(* IEC 61131-3 sources: rk/stdlib/generated, 8 files *)

(* ---- wasi-cli-types.st ---- *)
/* Generated from the WIT of wasi:cli@0.3.0. DO NOT EDIT! */
NAMESPACE INTERNAL Wasi
	NAMESPACE Cli
		NAMESPACE Types
			TYPE ERROR_CODE : USINT (
				IO := 0,
				ILLEGAL_BYTE_SEQUENCE := 1,
				PIPE := 2
			); END_TYPE
		END_NAMESPACE
	END_NAMESPACE
END_NAMESPACE

(* ---- wasi-clocks-system-clock.st ---- *)
/* Generated from the WIT of wasi:clocks@0.3.0. DO NOT EDIT! */
NAMESPACE INTERNAL Wasi
	NAMESPACE Clocks
		/* WASI System Clock is a clock API intended to let users query the current
		   time. The clock is not necessarily monotonic as it may be reset.

		   It is intended to be portable at least between Unix-family platforms and
		   Windows.

		   External references may be reset, so this clock is not necessarily
		   monotonic, making it unsuitable for measuring elapsed time.

		   It is intended for reporting the current date and time for humans. */
		NAMESPACE SystemClock
			/* An "instant", or "exact time", is a point in time without regard to any
			   time zone: just the time since a particular external reference point,
			   often called an "epoch".

			   Here, the epoch is 1970-01-01T00:00:00Z, also known as
			   [POSIX's Seconds Since the Epoch], also known as [Unix Time].

			   Note that even if the seconds field is negative, incrementing
			   nanoseconds always represents moving forwards in time.
			   For example, `{ -1 seconds, 999999999 nanoseconds }` represents the
			   instant one nanosecond before the epoch.
			   For more on various different ways to represent time, see
			   https://tc39.es/proposal-temporal/docs/timezone.html

			   [POSIX's Seconds Since the Epoch]: https://pubs.opengroup.org/onlinepubs/9699919799/xrat/V4_xbd_chap04.html#tag_21_04_16
			   [Unix Time]: https://en.wikipedia.org/wiki/Unix_time */
			TYPE INSTANT : STRUCT
				seconds : LINT;
				nanoseconds : UDINT;
			END_STRUCT END_TYPE

			/* `now` as the host gives it: the values of its result, which `NOW` puts
			   in its members. */
			{extern 'wasi:clocks/system-clock@0.3.0' 'now'}
			FUNCTION PRIVATE NOW_RAW
			VAR_OUTPUT
				seconds : LINT;
				nanoseconds : UDINT;
			END_VAR
			END_FUNCTION

			/* Read the current value of the clock.

			   This clock is not monotonic, therefore calling this function repeatedly
			   will not necessarily produce a sequence of non-decreasing values.

			   The nanoseconds field of the output is always less than 1000000000. */
			FUNCTION NOW : INSTANT
				NOW_RAW(seconds => NOW.seconds, nanoseconds => NOW.nanoseconds);
			END_FUNCTION

			/* Query the resolution of the clock. Returns the smallest duration of time
			   that the implementation permits distinguishing. */
			{extern 'wasi:clocks/system-clock@0.3.0' 'get-resolution'}
			FUNCTION GET_RESOLUTION : Wasi.Clocks.Types.DURATION
			END_FUNCTION
		END_NAMESPACE
	END_NAMESPACE
END_NAMESPACE

(* ---- wasi-clocks-types.st ---- *)
/* Generated from the WIT of wasi:clocks@0.3.0. DO NOT EDIT! */
NAMESPACE INTERNAL Wasi
	NAMESPACE Clocks
		/* This interface common types used throughout wasi:clocks. */
		NAMESPACE Types
			/* A duration of time, in nanoseconds. */
			TYPE DURATION : ULINT; END_TYPE
		END_NAMESPACE
	END_NAMESPACE
END_NAMESPACE

(* ---- wasi-clocks-timezone.st ---- *)
/* Generated from the WIT of wasi:clocks@0.3.0. DO NOT EDIT! */
NAMESPACE INTERNAL Wasi
	NAMESPACE Clocks
		NAMESPACE Timezone
			/* `iana-id` as the host gives it: its result in words of 8 bytes, as the
			   canonical ABI lays it out, which `IANA_ID` reads, and its string in
			   `value`, where the host writes it. */
			{extern 'wasi:clocks/timezone@0.3.0' 'iana-id'}
			FUNCTION PRIVATE IANA_ID_RAW
			VAR_IN_OUT
				value : STRING;
			END_VAR
			VAR_OUTPUT
				w0 : LWORD;
				w1 : LWORD;
			END_VAR
			END_FUNCTION

			/* Return the IANA identifier of the currently configured timezone. This
			   should be an identifier from the IANA Time Zone Database.

			   For displaying to a user, the identifier should be converted into a
			   localized name by means of an internationalization API.

			   If the implementation does not expose an actual timezone, or is unable
			   to provide mappings from times to deltas between the configured timezone
			   and UTC, or determining the current timezone fails, or the timezone does
			   not have an IANA identifier, this returns nothing. */
			FUNCTION IANA_ID
			VAR_IN_OUT
				value : STRING;
			END_VAR
			VAR_OUTPUT
				is_some : BOOL;
			END_VAR
			VAR
				w0 : LWORD;
				w1 : LWORD;
			END_VAR
				IANA_ID_RAW(value := value, w0 => w0, w1 => w1);
				is_some := w0.%X0;
			END_FUNCTION

			/* `utc-offset` as the host takes it: its parameters as the canonical ABI
			   passes them, which `UTC_OFFSET` passes field by field. */
			{extern 'wasi:clocks/timezone@0.3.0' 'utc-offset'}
			FUNCTION PRIVATE UTC_OFFSET_RAW
			VAR_INPUT
				when_seconds : LINT;
				when_nanoseconds : UDINT;
			END_VAR
			VAR_OUTPUT
				is_some : BOOL;
				value : LINT;
			END_VAR
			END_FUNCTION

			/* The number of nanoseconds difference between UTC time and the local
			   time of the currently configured timezone, at the exact time of
			   `instant`.

			   The magnitude of the returned value will always be less than
			   86,400,000,000,000 which is the number of nanoseconds in a day
			   (24*60*60*1e9).

			   If the implementation does not expose an actual timezone, or is unable
			   to provide mappings from times to deltas between the configured timezone
			   and UTC, or determining the current timezone fails, this returns
			   nothing. */
			FUNCTION UTC_OFFSET
			VAR_INPUT
				when : Wasi.Clocks.SystemClock.INSTANT;
			END_VAR
			VAR_OUTPUT
				is_some : BOOL;
				value : LINT;
			END_VAR
				UTC_OFFSET_RAW(when_seconds := when.seconds, when_nanoseconds := when.nanoseconds, is_some => is_some, value => value);
			END_FUNCTION

			/* `to-debug-string` as the host gives it: its result in words of 8 bytes,
			   as the canonical ABI lays it out, which `TO_DEBUG_STRING` reads, and its
			   string in `value`, where the host writes it. */
			{extern 'wasi:clocks/timezone@0.3.0' 'to-debug-string'}
			FUNCTION PRIVATE TO_DEBUG_STRING_RAW
			VAR_IN_OUT
				value : STRING;
			END_VAR
			VAR_OUTPUT
				w0 : LWORD;
				w1 : LWORD;
			END_VAR
			END_FUNCTION

			/* Returns a string that is suitable to assist humans in debugging whether
			   any timezone is available, and if so, which. This may be the same string
			   as `iana-id`, or a formatted representation of the UTC offset such as
			   `-04:00`, or something else.

			   WARNING: The returned string should not be consumed mechanically! It may
			   change across platforms, hosts, or other implementation details. Parsing
			   this string is a major platform-compatibility hazard. */
			FUNCTION TO_DEBUG_STRING
			VAR_IN_OUT
				value : STRING;
			END_VAR
			VAR
				w0 : LWORD;
				w1 : LWORD;
			END_VAR
				TO_DEBUG_STRING_RAW(value := value, w0 => w0, w1 => w1);
			END_FUNCTION
		END_NAMESPACE
	END_NAMESPACE
END_NAMESPACE

(* ---- wasi-cli-stderr.st ---- *)
/* Generated from the WIT of wasi:cli@0.3.0. DO NOT EDIT! */
NAMESPACE INTERNAL Wasi
	NAMESPACE Cli
		NAMESPACE Stderr
			/* Write the given stream to stderr.

			   If the stream's writable end is dropped this function will either return
			   success once the entire contents of the stream have been written or an
			   error-code representing a failure.

			   Otherwise if there is an error the readable end of the stream will be
			   dropped and this function will return an error-code. */
			{extern 'wasi:cli/stderr@0.3.0' 'write-via-stream'}
			FUNCTION WRITE_VIA_STREAM : UDINT
			VAR_INPUT
				data : UDINT;
			END_VAR
			END_FUNCTION

			/* Makes a stream of `u8`, and gives its reading end, then its writing end. */
			{extern 'wasi:cli/stderr@0.3.0' '[stream-new-0]write-via-stream'}
			FUNCTION BYTES_STREAM_NEW
			VAR_OUTPUT
				readable : UDINT;
				writable : UDINT;
			END_VAR
			END_FUNCTION

			/* Writes the bytes of `data`, as many as the reader takes: `written` of
			   them, after `DONE`. `closed` is TRUE once the reader has let go. */
			{extern async 'wasi:cli/stderr@0.3.0' '[stream-write-0]write-via-stream'}
			FUNCTION_BLOCK BYTES_STREAM_WRITE
			VAR_INPUT
				stream : UDINT;
				data : STRING[4096];
			END_VAR
			VAR_OUTPUT
				DONE : BOOL;
				written : UDINT;
				closed : BOOL;
			END_VAR
			END_FUNCTION_BLOCK

			/* Writes the `count` bytes from the one `data` points at, as many as the
			   reader takes: `written` of them, after `DONE`. The host reads them where
			   they are while the write runs, so they stay there, unchanged, until
			   `DONE`. `closed` is TRUE once the reader has let go. */
			{extern async 'wasi:cli/stderr@0.3.0' '[stream-write-0]write-via-stream'}
			FUNCTION_BLOCK BYTES_STREAM_WRITE_ARRAY
			VAR_INPUT
				stream : UDINT;
				data : REF_TO BYTE;
				count : UDINT;
			END_VAR
			VAR_OUTPUT
				DONE : BOOL;
				written : UDINT;
				closed : BOOL;
			END_VAR
			END_FUNCTION_BLOCK

			/* Lets go of the stream's reading end, `stream`. */
			{extern 'wasi:cli/stderr@0.3.0' '[stream-drop-readable-0]write-via-stream'}
			FUNCTION BYTES_STREAM_DROP_READABLE
			VAR_INPUT
				stream : UDINT;
			END_VAR
			END_FUNCTION

			/* Lets go of the stream's writing end, `stream`. */
			{extern 'wasi:cli/stderr@0.3.0' '[stream-drop-writable-0]write-via-stream'}
			FUNCTION BYTES_STREAM_DROP_WRITABLE
			VAR_INPUT
				stream : UDINT;
			END_VAR
			END_FUNCTION

			/* The bytes `IN` holds, which `BYTES_STREAM_WRITER` counts. */
			FUNCTION PRIVATE BYTES_STREAM_TEXT_LEN : UDINT
			VAR_INPUT
				IN : STRING[4096];
			END_VAR
				{wasm 'str.byte_len' (params IN) (result BYTES_STREAM_TEXT_LEN)}
			END_FUNCTION

			/* `IN` without its first `L` bytes: what `BYTES_STREAM_WRITER` has left to
			   write. */
			FUNCTION PRIVATE BYTES_STREAM_TEXT_AFTER : STRING[4096]
			VAR_INPUT
				IN : STRING[4096];
				L : UDINT;
			END_VAR
			VAR
				P : UDINT := 1;
			END_VAR
				{wasm 'str.byte_delete' (params IN L P) (result BYTES_STREAM_TEXT_AFTER)}
			END_FUNCTION

			/* Writes text to a stream of bytes it makes at its first call, for the
			   function `readable` is handed to. */
			FUNCTION_BLOCK BYTES_STREAM_WRITER
			VAR_INPUT
				/* A rising edge writes `IN`. An edge while `BUSY` is ignored. */
				REQ : BOOL;
				/* The text to write. */
				IN : STRING[4096];
				/* A rising edge ends the stream, once no write is under way. */
				CLOSE : BOOL;
			END_VAR
			VAR_OUTPUT
				/* The stream's reading end, to hand to the function that reads it. */
				readable : UDINT;
				/* TRUE while the reader has not taken all of `IN`. */
				BUSY : BOOL;
				/* TRUE in the call where the reader has taken all of `IN`, at once for an
				   empty text. */
				DONE : BOOL;
				/* TRUE once a write finds the reader gone, or a request comes after
				   `CLOSE`: the stream does not open again. */
				ERROR : BOOL;
			END_VAR
			VAR
				writable : UDINT;
				requested : BOOL;
				closing : BOOL;
				shut : BOOL;
				closed : BOOL;
				rest : STRING[4096];
				write : BYTES_STREAM_WRITE;
			END_VAR
			VAR_TEMP
				again : BOOL;
			END_VAR
				IF writable = 0 AND NOT closed THEN
					BYTES_STREAM_NEW(readable => readable, writable => writable);
				END_IF;
				DONE := FALSE;
				// An edge while BUSY is ignored.
				IF REQ AND NOT requested AND NOT BUSY THEN
					ERROR := closed;
					IF NOT closed THEN
						// A write of no bytes asks the reader whether it is ready,
						// which it may answer late: an empty text is done here.
						IF BYTES_STREAM_TEXT_LEN(IN) = 0 THEN
							DONE := TRUE;
						ELSE
							rest := IN;
							BUSY := TRUE;
						END_IF;
					END_IF;
				END_IF;
				requested := REQ;
				IF BUSY THEN
					// Each pass after the first hands over a byte at least, so the
					// loop ends.
					REPEAT
						again := FALSE;
						// Starts the write of the rest, or checks the one running.
						write(stream := writable, data := rest);
						IF write.DONE THEN
							IF write.closed THEN
								// The reader left: the writing end goes too.
								BYTES_STREAM_DROP_WRITABLE(stream := writable);
								writable := 0;
								closed := TRUE;
								BUSY := FALSE;
								ERROR := TRUE;
							ELSIF write.written < BYTES_STREAM_TEXT_LEN(rest) THEN
								// The reader took a part: the rest goes next, at once while
								// it takes some.
								rest := BYTES_STREAM_TEXT_AFTER(rest, write.written);
								again := write.written > 0;
							ELSE
								BUSY := FALSE;
								DONE := TRUE;
							END_IF;
						END_IF;
					UNTIL NOT again
					END_REPEAT;
				END_IF;
				// The writing end goes once no write is under way.
				IF CLOSE AND NOT closing THEN
					shut := TRUE;
				END_IF;
				closing := CLOSE;
				IF shut AND NOT BUSY THEN
					IF writable <> 0 THEN
						BYTES_STREAM_DROP_WRITABLE(stream := writable);
						writable := 0;
					END_IF;
					closed := TRUE;
					shut := FALSE;
				END_IF;
			END_FUNCTION_BLOCK

			/* The subscript of the first byte of `IN`, which
			   `BYTES_STREAM_ARRAY_WRITER` writes from. */
			FUNCTION PRIVATE BYTES_STREAM_ARRAY_FIRST : LINT
			VAR_INPUT
				IN : ARRAY[*] OF BYTE;
			END_VAR
			VAR
				DIM : DINT := 1;
			END_VAR
				{wasm 'array.lower_bound' (params IN DIM) (result BYTES_STREAM_ARRAY_FIRST)}
			END_FUNCTION

			/* How many bytes `IN` holds, which `BYTES_STREAM_ARRAY_WRITER` writes at
			   most. */
			FUNCTION PRIVATE BYTES_STREAM_ARRAY_LEN : LINT
			VAR_INPUT
				IN : ARRAY[*] OF BYTE;
			END_VAR
			VAR
				DIM : DINT := 1;
				lower : LINT;
				upper : LINT;
			END_VAR
				{wasm 'array.lower_bound' (params IN DIM) (result lower)}
				{wasm 'array.upper_bound' (params IN DIM) (result upper)}
				BYTES_STREAM_ARRAY_LEN := upper - lower + 1;
			END_FUNCTION

			/* Writes bytes from an array to a stream of bytes it makes at its first
			   call, for the function `readable` is handed to. */
			FUNCTION_BLOCK BYTES_STREAM_ARRAY_WRITER
			VAR_INPUT
				/* A rising edge writes the first `COUNT` bytes of `IN`. An edge while
				   `BUSY` is ignored. */
				REQ : BOOL;
				/* How many bytes of `IN` a request writes, from its first on. */
				COUNT : UDINT;
				/* A rising edge ends the stream, once no write is under way. */
				CLOSE : BOOL;
			END_VAR
			VAR_IN_OUT
				/* The bytes to write. The host reads them where they are while `BUSY`:
				   they stay as they are until `DONE`. */
				IN : ARRAY[*] OF BYTE;
			END_VAR
			VAR_OUTPUT
				/* The stream's reading end, to hand to the function that reads it. */
				readable : UDINT;
				/* TRUE while the reader has not taken all `COUNT` bytes. */
				BUSY : BOOL;
				/* TRUE in the call where the reader has taken all `COUNT` bytes, at once
				   for none. */
				DONE : BOOL;
				/* TRUE once a write finds the reader gone, or a request comes after
				   `CLOSE`: the stream does not open again. */
				ERROR : BOOL;
			END_VAR
			VAR
				writable : UDINT;
				requested : BOOL;
				closing : BOOL;
				shut : BOOL;
				closed : BOOL;
				total : UDINT;
				sent : UDINT;
				base : LINT;
				write : BYTES_STREAM_WRITE_ARRAY;
			END_VAR
			VAR_TEMP
				again : BOOL;
				offset : LINT;
			END_VAR
				IF writable = 0 AND NOT closed THEN
					BYTES_STREAM_NEW(readable => readable, writable => writable);
				END_IF;
				DONE := FALSE;
				// An edge while BUSY is ignored.
				IF REQ AND NOT requested AND NOT BUSY THEN
					ERROR := closed;
					IF NOT closed THEN
						// A write of no bytes asks the reader whether it is ready,
						// which it may answer late: none is done here.
						IF COUNT = 0 THEN
							DONE := TRUE;
						ELSIF COUNT > BYTES_STREAM_ARRAY_LEN(IN) THEN
							__RAISE('COUNT is past the end of IN');
						ELSE
							total := COUNT;
							sent := 0;
							base := BYTES_STREAM_ARRAY_FIRST(IN);
							BUSY := TRUE;
						END_IF;
					END_IF;
				END_IF;
				requested := REQ;
				IF BUSY THEN
					// Each pass after the first hands over a byte at least, so the
					// loop ends.
					REPEAT
						again := FALSE;
						offset := sent;
						// Starts the write of the bytes not taken yet, from where they
						// are, or checks the one running.
						write(stream := writable, data := REF(IN[base + offset]), count := total - sent);
						IF write.DONE THEN
							IF write.closed THEN
								// The reader left: the writing end goes too.
								BYTES_STREAM_DROP_WRITABLE(stream := writable);
								writable := 0;
								closed := TRUE;
								BUSY := FALSE;
								ERROR := TRUE;
							ELSIF write.written < total - sent THEN
								// The reader took a part: the rest goes next, at once while
								// it takes some.
								sent := sent + write.written;
								again := write.written > 0;
							ELSE
								BUSY := FALSE;
								DONE := TRUE;
							END_IF;
						END_IF;
					UNTIL NOT again
					END_REPEAT;
				END_IF;
				// The writing end goes once no write is under way.
				IF CLOSE AND NOT closing THEN
					shut := TRUE;
				END_IF;
				closing := CLOSE;
				IF shut AND NOT BUSY THEN
					IF writable <> 0 THEN
						BYTES_STREAM_DROP_WRITABLE(stream := writable);
						writable := 0;
					END_IF;
					closed := TRUE;
					shut := FALSE;
				END_IF;
			END_FUNCTION_BLOCK

			/* Reads the value the future holds, which comes back after `DONE`. */
			{extern async 'wasi:cli/stderr@0.3.0' '[future-read-1]write-via-stream'}
			FUNCTION_BLOCK RESULT_FUTURE_READ
			VAR_INPUT
				future : UDINT;
			END_VAR
			VAR_OUTPUT
				DONE : BOOL;
				failed : BOOL;
				error : Wasi.Cli.Types.ERROR_CODE;
			END_VAR
			END_FUNCTION_BLOCK

			/* Lets go of the future's reading end, `future`. */
			{extern 'wasi:cli/stderr@0.3.0' '[future-drop-readable-1]write-via-stream'}
			FUNCTION RESULT_FUTURE_DROP_READABLE
			VAR_INPUT
				future : UDINT;
			END_VAR
			END_FUNCTION

			/* Reads the value the future holds, which comes back after `DONE`, then
			   lets go of the future's reading end: `future` is 0 from then on, and a
			   call with `future` 0 does nothing. */
			FUNCTION_BLOCK RESULT_FUTURE_GET
			VAR_IN_OUT
				future : UDINT;
			END_VAR
			VAR_OUTPUT
				DONE : BOOL;
				failed : BOOL;
				error : Wasi.Cli.Types.ERROR_CODE;
			END_VAR
			VAR
				call : RESULT_FUTURE_READ;
			END_VAR
				DONE := FALSE;
				IF future <> 0 THEN
					call(future := future);
					IF call.DONE THEN
						failed := call.failed;
						error := call.error;
						RESULT_FUTURE_DROP_READABLE(future := future);
						future := 0;
						DONE := TRUE;
					END_IF;
				END_IF;
			END_FUNCTION_BLOCK

			/* Writes text to `write-via-stream` through a stream of bytes it opens at
			   the first request. */
			FUNCTION_BLOCK WRITE_VIA_STREAM_WRITER
			VAR_INPUT
				/* A rising edge writes `IN`; the first opens the stream and calls
				   `write-via-stream` with it. An edge while `BUSY` is ignored. */
				REQ : BOOL;
				/* The text to write. */
				IN : STRING[4096];
				/* A rising edge ends the stream, once no write is under way. */
				CLOSE : BOOL;
			END_VAR
			VAR_OUTPUT
				/* TRUE while the reader has not taken all of `IN`. */
				BUSY : BOOL;
				/* TRUE in the call where the reader has taken all of `IN`, at once for an
				   empty text. */
				DONE : BOOL;
				/* TRUE once a write finds the reader gone, a request comes after `CLOSE`,
				   or the `result<_, error-code>` from `write-via-stream` is an error,
				   whose `error-code` is in `ERRORID`. */
				ERROR : BOOL;
				/* The `error-code` of the `result<_, error-code>` from `write-via-stream`,
				   when it is an error, which turns `ERROR` TRUE. */
				ERRORID : Wasi.Cli.Types.ERROR_CODE;
				/* TRUE once the `future<result<_, error-code>>` from `write-via-stream`
				   has its value. */
				ENDED : BOOL;
			END_VAR
			VAR
				open : BOOL;
				stream : BYTES_STREAM_WRITER;
				future : UDINT;
				answer : RESULT_FUTURE_GET;
			END_VAR
				// The stream, made at the first request and handed to the function.
				IF REQ AND NOT open THEN
					stream(REQ := FALSE, IN := IN, CLOSE := FALSE);
					future := Wasi.Cli.Stderr.WRITE_VIA_STREAM(data := stream.readable);
					open := TRUE;
				END_IF;
				IF open THEN
					stream(REQ := REQ, IN := IN, CLOSE := CLOSE);
					BUSY := stream.BUSY;
					DONE := stream.DONE;
					// The answer, read once it comes, and kept.
					answer(future := future);
					IF answer.DONE THEN
						ERRORID := answer.error;
						ENDED := TRUE;
					END_IF;
					ERROR := stream.ERROR OR answer.failed;
				END_IF;
			END_FUNCTION_BLOCK

			/* Writes bytes from an array to `write-via-stream` through a stream of
			   bytes it opens at the first request. */
			FUNCTION_BLOCK WRITE_VIA_STREAM_ARRAY_WRITER
			VAR_INPUT
				/* A rising edge writes the first `COUNT` bytes of `IN`; the first opens
				   the stream and calls `write-via-stream` with it. An edge while `BUSY` is
				   ignored. */
				REQ : BOOL;
				/* How many bytes of `IN` a request writes, from its first on. */
				COUNT : UDINT;
				/* A rising edge ends the stream, once no write is under way. */
				CLOSE : BOOL;
			END_VAR
			VAR_IN_OUT
				/* The bytes to write. The host reads them where they are while `BUSY`:
				   they stay as they are until `DONE`. */
				IN : ARRAY[*] OF BYTE;
			END_VAR
			VAR_OUTPUT
				/* TRUE while the reader has not taken all `COUNT` bytes. */
				BUSY : BOOL;
				/* TRUE in the call where the reader has taken all `COUNT` bytes, at once
				   for none. */
				DONE : BOOL;
				/* TRUE once a write finds the reader gone, a request comes after `CLOSE`,
				   or the `result<_, error-code>` from `write-via-stream` is an error,
				   whose `error-code` is in `ERRORID`. */
				ERROR : BOOL;
				/* The `error-code` of the `result<_, error-code>` from `write-via-stream`,
				   when it is an error, which turns `ERROR` TRUE. */
				ERRORID : Wasi.Cli.Types.ERROR_CODE;
				/* TRUE once the `future<result<_, error-code>>` from `write-via-stream`
				   has its value. */
				ENDED : BOOL;
			END_VAR
			VAR
				open : BOOL;
				stream : BYTES_STREAM_ARRAY_WRITER;
				future : UDINT;
				answer : RESULT_FUTURE_GET;
			END_VAR
				// The stream, made at the first request and handed to the function.
				IF REQ AND NOT open THEN
					stream(REQ := FALSE, COUNT := COUNT, CLOSE := FALSE, IN := IN);
					future := Wasi.Cli.Stderr.WRITE_VIA_STREAM(data := stream.readable);
					open := TRUE;
				END_IF;
				IF open THEN
					stream(REQ := REQ, COUNT := COUNT, CLOSE := CLOSE, IN := IN);
					BUSY := stream.BUSY;
					DONE := stream.DONE;
					// The answer, read once it comes, and kept.
					answer(future := future);
					IF answer.DONE THEN
						ERRORID := answer.error;
						ENDED := TRUE;
					END_IF;
					ERROR := stream.ERROR OR answer.failed;
				END_IF;
			END_FUNCTION_BLOCK
		END_NAMESPACE
	END_NAMESPACE
END_NAMESPACE
/* Not generated:
   - `BYTES_STREAM_CANCEL_WRITE`: a cancel blocks the scan.
   - `RESULT_FUTURE_CANCEL_READ`: a cancel blocks the scan. */

(* ---- wasi-cli-stdin.st ---- *)
/* Generated from the WIT of wasi:cli@0.3.0. DO NOT EDIT! */
NAMESPACE INTERNAL Wasi
	NAMESPACE Cli
		NAMESPACE Stdin
			/* Return a stream for reading from stdin.

			   This function returns a stream which provides data read from stdin,
			   and a future to signal read results.

			   If the stream's readable end is dropped the future will resolve to success.

			   If the stream's writable end is dropped the future will either resolve to
			   success if stdin was closed by the writer or to an error-code if reading
			   failed for some other reason.

			   Multiple streams may be active at the same time. The behavior of concurrent
			   reads is implementation-specific. */
			{extern 'wasi:cli/stdin@0.3.0' 'read-via-stream'}
			FUNCTION READ_VIA_STREAM
			VAR_OUTPUT
				item0 : UDINT;
				item1 : UDINT;
			END_VAR
			END_FUNCTION

			/* Reads the bytes that come next into `data`, as many as it holds at most:
			   `read` of them, after `DONE`. `closed` is TRUE once the writer has let
			   go. */
			{extern async 'wasi:cli/stdin@0.3.0' '[stream-read-0]read-via-stream'}
			FUNCTION_BLOCK BYTES_STREAM_READ
			VAR_INPUT
				stream : UDINT;
			END_VAR
			VAR_OUTPUT
				DONE : BOOL;
				data : STRING[4096];
				read : UDINT;
				closed : BOOL;
			END_VAR
			END_FUNCTION_BLOCK

			/* Reads the bytes that come next into `data`, as many as it holds at most:
			   `read` of them, after `DONE`. `closed` is TRUE once the writer has let
			   go. */
			{extern async 'wasi:cli/stdin@0.3.0' '[stream-read-0]read-via-stream'}
			FUNCTION_BLOCK BYTES_STREAM_READ_ARRAY
			VAR_INPUT
				stream : UDINT;
			END_VAR
			VAR_OUTPUT
				DONE : BOOL;
				data : ARRAY[0..8191] OF BYTE;
				read : UDINT;
				closed : BOOL;
			END_VAR
			END_FUNCTION_BLOCK

			/* Lets go of the stream's reading end, `stream`. */
			{extern 'wasi:cli/stdin@0.3.0' '[stream-drop-readable-0]read-via-stream'}
			FUNCTION BYTES_STREAM_DROP_READABLE
			VAR_INPUT
				stream : UDINT;
			END_VAR
			END_FUNCTION

			/* Reads the value the future holds, which comes back after `DONE`. */
			{extern async 'wasi:cli/stdin@0.3.0' '[future-read-1]read-via-stream'}
			FUNCTION_BLOCK RESULT_FUTURE_READ
			VAR_INPUT
				future : UDINT;
			END_VAR
			VAR_OUTPUT
				DONE : BOOL;
				failed : BOOL;
				error : Wasi.Cli.Types.ERROR_CODE;
			END_VAR
			END_FUNCTION_BLOCK

			/* Lets go of the future's reading end, `future`. */
			{extern 'wasi:cli/stdin@0.3.0' '[future-drop-readable-1]read-via-stream'}
			FUNCTION RESULT_FUTURE_DROP_READABLE
			VAR_INPUT
				future : UDINT;
			END_VAR
			END_FUNCTION

			/* Reads the value the future holds, which comes back after `DONE`, then
			   lets go of the future's reading end: `future` is 0 from then on, and a
			   call with `future` 0 does nothing. */
			FUNCTION_BLOCK RESULT_FUTURE_GET
			VAR_IN_OUT
				future : UDINT;
			END_VAR
			VAR_OUTPUT
				DONE : BOOL;
				failed : BOOL;
				error : Wasi.Cli.Types.ERROR_CODE;
			END_VAR
			VAR
				call : RESULT_FUTURE_READ;
			END_VAR
				DONE := FALSE;
				IF future <> 0 THEN
					call(future := future);
					IF call.DONE THEN
						failed := call.failed;
						error := call.error;
						RESULT_FUTURE_DROP_READABLE(future := future);
						future := 0;
						DONE := TRUE;
					END_IF;
				END_IF;
			END_FUNCTION_BLOCK

			/* Reads what `read-via-stream` gives through a stream of bytes, a request
			   at a time. */
			FUNCTION_BLOCK READ_VIA_STREAM_READER
			VAR_INPUT
				/* A rising edge reads what comes next, 4096 bytes at most; the first calls
				   `read-via-stream`. An edge while `BUSY` is ignored, and one after the
				   stream ended is `DONE` at once, `OUT` empty. */
				REQ : BOOL;
				/* A rising edge lets go of the stream, once no read is under way. */
				CLOSE : BOOL;
			END_VAR
			VAR_OUTPUT
				/* TRUE while a read waits for bytes. */
				BUSY : BOOL;
				/* TRUE in the call where a read has given what came, in `OUT`. */
				DONE : BOOL;
				/* What the last read gave: empty once the stream has ended, nothing more
				   coming. */
				OUT : STRING[4096];
				/* TRUE once the `result<_, error-code>` from `read-via-stream` is an
				   error, whose `error-code` is in `ERRORID`. */
				ERROR : BOOL;
				/* The `error-code` of the `result<_, error-code>` from `read-via-stream`,
				   when it is an error, which turns `ERROR` TRUE. */
				ERRORID : Wasi.Cli.Types.ERROR_CODE;
				/* TRUE once the stream has ended and the `future<result<_, error-code>>`
				   from `read-via-stream` has its value. */
				ENDED : BOOL;
			END_VAR
			VAR
				open : BOOL;
				requested : BOOL;
				closing : BOOL;
				shut : BOOL;
				stream : UDINT;
				future : UDINT;
				read : BYTES_STREAM_READ;
				answer : RESULT_FUTURE_GET;
				came : BOOL;
			END_VAR
				DONE := FALSE;
				// The stream, given by the function at the first request.
				IF REQ AND NOT open THEN
					Wasi.Cli.Stdin.READ_VIA_STREAM(item0 => stream, item1 => future);
					open := TRUE;
				END_IF;
				IF open THEN
					// An edge while BUSY is ignored.
					IF REQ AND NOT requested AND NOT BUSY THEN
						IF stream <> 0 THEN
							BUSY := TRUE;
						ELSE
							// The stream has ended: nothing more comes.
							OUT := '';
							DONE := TRUE;
						END_IF;
					END_IF;
					requested := REQ;
					IF BUSY THEN
						// Starts the read, or checks the one running.
						read(stream := stream);
						IF read.DONE THEN
							OUT := read.data;
							BUSY := FALSE;
							DONE := TRUE;
							IF read.closed THEN
								// The writer left: the reading end goes too.
								BYTES_STREAM_DROP_READABLE(stream := stream);
								stream := 0;
							END_IF;
						END_IF;
					END_IF;
					// The reading end goes on CLOSE, once no read is under way.
					IF CLOSE AND NOT closing THEN
						shut := TRUE;
					END_IF;
					closing := CLOSE;
					IF shut AND NOT BUSY THEN
						IF stream <> 0 THEN
							BYTES_STREAM_DROP_READABLE(stream := stream);
							stream := 0;
						END_IF;
						shut := FALSE;
					END_IF;
					// The answer, read once it comes, and kept.
					answer(future := future);
					IF answer.DONE THEN
						ERRORID := answer.error;
						came := TRUE;
					END_IF;
					ENDED := stream = 0 AND came;
					ERROR := answer.failed;
				END_IF;
			END_FUNCTION_BLOCK

			/* Reads what `read-via-stream` gives through a stream of bytes into an
			   array, a request at a time. */
			FUNCTION_BLOCK READ_VIA_STREAM_ARRAY_READER
			VAR_INPUT
				/* A rising edge reads what comes next, 8192 bytes at most; the first calls
				   `read-via-stream`. An edge while `BUSY` is ignored, and one after the
				   stream ended is `DONE` at once, `COUNT` 0. */
				REQ : BOOL;
				/* A rising edge lets go of the stream, once no read is under way. */
				CLOSE : BOOL;
			END_VAR
			VAR_OUTPUT
				/* TRUE while a read waits for bytes. */
				BUSY : BOOL;
				/* TRUE in the call where a read has given what came, in `OUT`. */
				DONE : BOOL;
				/* The bytes the last read gave, its first `COUNT`. */
				OUT : ARRAY[0..8191] OF BYTE;
				/* How many bytes the last read gave: 0 once the stream has ended, nothing
				   more coming. */
				COUNT : UDINT;
				/* TRUE once the `result<_, error-code>` from `read-via-stream` is an
				   error, whose `error-code` is in `ERRORID`. */
				ERROR : BOOL;
				/* The `error-code` of the `result<_, error-code>` from `read-via-stream`,
				   when it is an error, which turns `ERROR` TRUE. */
				ERRORID : Wasi.Cli.Types.ERROR_CODE;
				/* TRUE once the stream has ended and the `future<result<_, error-code>>`
				   from `read-via-stream` has its value. */
				ENDED : BOOL;
			END_VAR
			VAR
				open : BOOL;
				requested : BOOL;
				closing : BOOL;
				shut : BOOL;
				stream : UDINT;
				future : UDINT;
				read : BYTES_STREAM_READ_ARRAY;
				answer : RESULT_FUTURE_GET;
				came : BOOL;
			END_VAR
				DONE := FALSE;
				// The stream, given by the function at the first request.
				IF REQ AND NOT open THEN
					Wasi.Cli.Stdin.READ_VIA_STREAM(item0 => stream, item1 => future);
					open := TRUE;
				END_IF;
				IF open THEN
					// An edge while BUSY is ignored.
					IF REQ AND NOT requested AND NOT BUSY THEN
						IF stream <> 0 THEN
							BUSY := TRUE;
						ELSE
							// The stream has ended: nothing more comes.
							COUNT := 0;
							DONE := TRUE;
						END_IF;
					END_IF;
					requested := REQ;
					IF BUSY THEN
						// Starts the read, or checks the one running.
						read(stream := stream);
						IF read.DONE THEN
							OUT := read.data;
							COUNT := read.read;
							BUSY := FALSE;
							DONE := TRUE;
							IF read.closed THEN
								// The writer left: the reading end goes too.
								BYTES_STREAM_DROP_READABLE(stream := stream);
								stream := 0;
							END_IF;
						END_IF;
					END_IF;
					// The reading end goes on CLOSE, once no read is under way.
					IF CLOSE AND NOT closing THEN
						shut := TRUE;
					END_IF;
					closing := CLOSE;
					IF shut AND NOT BUSY THEN
						IF stream <> 0 THEN
							BYTES_STREAM_DROP_READABLE(stream := stream);
							stream := 0;
						END_IF;
						shut := FALSE;
					END_IF;
					// The answer, read once it comes, and kept.
					answer(future := future);
					IF answer.DONE THEN
						ERRORID := answer.error;
						came := TRUE;
					END_IF;
					ENDED := stream = 0 AND came;
					ERROR := answer.failed;
				END_IF;
			END_FUNCTION_BLOCK
		END_NAMESPACE
	END_NAMESPACE
END_NAMESPACE
/* Not generated:
   - `BYTES_STREAM_CANCEL_READ`: a cancel blocks the scan.
   - `RESULT_FUTURE_CANCEL_READ`: a cancel blocks the scan. */

(* ---- wasi-cli-stdout.st ---- *)
/* Generated from the WIT of wasi:cli@0.3.0. DO NOT EDIT! */
NAMESPACE INTERNAL Wasi
	NAMESPACE Cli
		NAMESPACE Stdout
			/* Write the given stream to stdout.

			   If the stream's writable end is dropped this function will either return
			   success once the entire contents of the stream have been written or an
			   error-code representing a failure.

			   Otherwise if there is an error the readable end of the stream will be
			   dropped and this function will return an error-code. */
			{extern 'wasi:cli/stdout@0.3.0' 'write-via-stream'}
			FUNCTION WRITE_VIA_STREAM : UDINT
			VAR_INPUT
				data : UDINT;
			END_VAR
			END_FUNCTION

			/* Makes a stream of `u8`, and gives its reading end, then its writing end. */
			{extern 'wasi:cli/stdout@0.3.0' '[stream-new-0]write-via-stream'}
			FUNCTION BYTES_STREAM_NEW
			VAR_OUTPUT
				readable : UDINT;
				writable : UDINT;
			END_VAR
			END_FUNCTION

			/* Writes the bytes of `data`, as many as the reader takes: `written` of
			   them, after `DONE`. `closed` is TRUE once the reader has let go. */
			{extern async 'wasi:cli/stdout@0.3.0' '[stream-write-0]write-via-stream'}
			FUNCTION_BLOCK BYTES_STREAM_WRITE
			VAR_INPUT
				stream : UDINT;
				data : STRING[4096];
			END_VAR
			VAR_OUTPUT
				DONE : BOOL;
				written : UDINT;
				closed : BOOL;
			END_VAR
			END_FUNCTION_BLOCK

			/* Writes the `count` bytes from the one `data` points at, as many as the
			   reader takes: `written` of them, after `DONE`. The host reads them where
			   they are while the write runs, so they stay there, unchanged, until
			   `DONE`. `closed` is TRUE once the reader has let go. */
			{extern async 'wasi:cli/stdout@0.3.0' '[stream-write-0]write-via-stream'}
			FUNCTION_BLOCK BYTES_STREAM_WRITE_ARRAY
			VAR_INPUT
				stream : UDINT;
				data : REF_TO BYTE;
				count : UDINT;
			END_VAR
			VAR_OUTPUT
				DONE : BOOL;
				written : UDINT;
				closed : BOOL;
			END_VAR
			END_FUNCTION_BLOCK

			/* Lets go of the stream's reading end, `stream`. */
			{extern 'wasi:cli/stdout@0.3.0' '[stream-drop-readable-0]write-via-stream'}
			FUNCTION BYTES_STREAM_DROP_READABLE
			VAR_INPUT
				stream : UDINT;
			END_VAR
			END_FUNCTION

			/* Lets go of the stream's writing end, `stream`. */
			{extern 'wasi:cli/stdout@0.3.0' '[stream-drop-writable-0]write-via-stream'}
			FUNCTION BYTES_STREAM_DROP_WRITABLE
			VAR_INPUT
				stream : UDINT;
			END_VAR
			END_FUNCTION

			/* The bytes `IN` holds, which `BYTES_STREAM_WRITER` counts. */
			FUNCTION PRIVATE BYTES_STREAM_TEXT_LEN : UDINT
			VAR_INPUT
				IN : STRING[4096];
			END_VAR
				{wasm 'str.byte_len' (params IN) (result BYTES_STREAM_TEXT_LEN)}
			END_FUNCTION

			/* `IN` without its first `L` bytes: what `BYTES_STREAM_WRITER` has left to
			   write. */
			FUNCTION PRIVATE BYTES_STREAM_TEXT_AFTER : STRING[4096]
			VAR_INPUT
				IN : STRING[4096];
				L : UDINT;
			END_VAR
			VAR
				P : UDINT := 1;
			END_VAR
				{wasm 'str.byte_delete' (params IN L P) (result BYTES_STREAM_TEXT_AFTER)}
			END_FUNCTION

			/* Writes text to a stream of bytes it makes at its first call, for the
			   function `readable` is handed to. */
			FUNCTION_BLOCK BYTES_STREAM_WRITER
			VAR_INPUT
				/* A rising edge writes `IN`. An edge while `BUSY` is ignored. */
				REQ : BOOL;
				/* The text to write. */
				IN : STRING[4096];
				/* A rising edge ends the stream, once no write is under way. */
				CLOSE : BOOL;
			END_VAR
			VAR_OUTPUT
				/* The stream's reading end, to hand to the function that reads it. */
				readable : UDINT;
				/* TRUE while the reader has not taken all of `IN`. */
				BUSY : BOOL;
				/* TRUE in the call where the reader has taken all of `IN`, at once for an
				   empty text. */
				DONE : BOOL;
				/* TRUE once a write finds the reader gone, or a request comes after
				   `CLOSE`: the stream does not open again. */
				ERROR : BOOL;
			END_VAR
			VAR
				writable : UDINT;
				requested : BOOL;
				closing : BOOL;
				shut : BOOL;
				closed : BOOL;
				rest : STRING[4096];
				write : BYTES_STREAM_WRITE;
			END_VAR
			VAR_TEMP
				again : BOOL;
			END_VAR
				IF writable = 0 AND NOT closed THEN
					BYTES_STREAM_NEW(readable => readable, writable => writable);
				END_IF;
				DONE := FALSE;
				// An edge while BUSY is ignored.
				IF REQ AND NOT requested AND NOT BUSY THEN
					ERROR := closed;
					IF NOT closed THEN
						// A write of no bytes asks the reader whether it is ready,
						// which it may answer late: an empty text is done here.
						IF BYTES_STREAM_TEXT_LEN(IN) = 0 THEN
							DONE := TRUE;
						ELSE
							rest := IN;
							BUSY := TRUE;
						END_IF;
					END_IF;
				END_IF;
				requested := REQ;
				IF BUSY THEN
					// Each pass after the first hands over a byte at least, so the
					// loop ends.
					REPEAT
						again := FALSE;
						// Starts the write of the rest, or checks the one running.
						write(stream := writable, data := rest);
						IF write.DONE THEN
							IF write.closed THEN
								// The reader left: the writing end goes too.
								BYTES_STREAM_DROP_WRITABLE(stream := writable);
								writable := 0;
								closed := TRUE;
								BUSY := FALSE;
								ERROR := TRUE;
							ELSIF write.written < BYTES_STREAM_TEXT_LEN(rest) THEN
								// The reader took a part: the rest goes next, at once while
								// it takes some.
								rest := BYTES_STREAM_TEXT_AFTER(rest, write.written);
								again := write.written > 0;
							ELSE
								BUSY := FALSE;
								DONE := TRUE;
							END_IF;
						END_IF;
					UNTIL NOT again
					END_REPEAT;
				END_IF;
				// The writing end goes once no write is under way.
				IF CLOSE AND NOT closing THEN
					shut := TRUE;
				END_IF;
				closing := CLOSE;
				IF shut AND NOT BUSY THEN
					IF writable <> 0 THEN
						BYTES_STREAM_DROP_WRITABLE(stream := writable);
						writable := 0;
					END_IF;
					closed := TRUE;
					shut := FALSE;
				END_IF;
			END_FUNCTION_BLOCK

			/* The subscript of the first byte of `IN`, which
			   `BYTES_STREAM_ARRAY_WRITER` writes from. */
			FUNCTION PRIVATE BYTES_STREAM_ARRAY_FIRST : LINT
			VAR_INPUT
				IN : ARRAY[*] OF BYTE;
			END_VAR
			VAR
				DIM : DINT := 1;
			END_VAR
				{wasm 'array.lower_bound' (params IN DIM) (result BYTES_STREAM_ARRAY_FIRST)}
			END_FUNCTION

			/* How many bytes `IN` holds, which `BYTES_STREAM_ARRAY_WRITER` writes at
			   most. */
			FUNCTION PRIVATE BYTES_STREAM_ARRAY_LEN : LINT
			VAR_INPUT
				IN : ARRAY[*] OF BYTE;
			END_VAR
			VAR
				DIM : DINT := 1;
				lower : LINT;
				upper : LINT;
			END_VAR
				{wasm 'array.lower_bound' (params IN DIM) (result lower)}
				{wasm 'array.upper_bound' (params IN DIM) (result upper)}
				BYTES_STREAM_ARRAY_LEN := upper - lower + 1;
			END_FUNCTION

			/* Writes bytes from an array to a stream of bytes it makes at its first
			   call, for the function `readable` is handed to. */
			FUNCTION_BLOCK BYTES_STREAM_ARRAY_WRITER
			VAR_INPUT
				/* A rising edge writes the first `COUNT` bytes of `IN`. An edge while
				   `BUSY` is ignored. */
				REQ : BOOL;
				/* How many bytes of `IN` a request writes, from its first on. */
				COUNT : UDINT;
				/* A rising edge ends the stream, once no write is under way. */
				CLOSE : BOOL;
			END_VAR
			VAR_IN_OUT
				/* The bytes to write. The host reads them where they are while `BUSY`:
				   they stay as they are until `DONE`. */
				IN : ARRAY[*] OF BYTE;
			END_VAR
			VAR_OUTPUT
				/* The stream's reading end, to hand to the function that reads it. */
				readable : UDINT;
				/* TRUE while the reader has not taken all `COUNT` bytes. */
				BUSY : BOOL;
				/* TRUE in the call where the reader has taken all `COUNT` bytes, at once
				   for none. */
				DONE : BOOL;
				/* TRUE once a write finds the reader gone, or a request comes after
				   `CLOSE`: the stream does not open again. */
				ERROR : BOOL;
			END_VAR
			VAR
				writable : UDINT;
				requested : BOOL;
				closing : BOOL;
				shut : BOOL;
				closed : BOOL;
				total : UDINT;
				sent : UDINT;
				base : LINT;
				write : BYTES_STREAM_WRITE_ARRAY;
			END_VAR
			VAR_TEMP
				again : BOOL;
				offset : LINT;
			END_VAR
				IF writable = 0 AND NOT closed THEN
					BYTES_STREAM_NEW(readable => readable, writable => writable);
				END_IF;
				DONE := FALSE;
				// An edge while BUSY is ignored.
				IF REQ AND NOT requested AND NOT BUSY THEN
					ERROR := closed;
					IF NOT closed THEN
						// A write of no bytes asks the reader whether it is ready,
						// which it may answer late: none is done here.
						IF COUNT = 0 THEN
							DONE := TRUE;
						ELSIF COUNT > BYTES_STREAM_ARRAY_LEN(IN) THEN
							__RAISE('COUNT is past the end of IN');
						ELSE
							total := COUNT;
							sent := 0;
							base := BYTES_STREAM_ARRAY_FIRST(IN);
							BUSY := TRUE;
						END_IF;
					END_IF;
				END_IF;
				requested := REQ;
				IF BUSY THEN
					// Each pass after the first hands over a byte at least, so the
					// loop ends.
					REPEAT
						again := FALSE;
						offset := sent;
						// Starts the write of the bytes not taken yet, from where they
						// are, or checks the one running.
						write(stream := writable, data := REF(IN[base + offset]), count := total - sent);
						IF write.DONE THEN
							IF write.closed THEN
								// The reader left: the writing end goes too.
								BYTES_STREAM_DROP_WRITABLE(stream := writable);
								writable := 0;
								closed := TRUE;
								BUSY := FALSE;
								ERROR := TRUE;
							ELSIF write.written < total - sent THEN
								// The reader took a part: the rest goes next, at once while
								// it takes some.
								sent := sent + write.written;
								again := write.written > 0;
							ELSE
								BUSY := FALSE;
								DONE := TRUE;
							END_IF;
						END_IF;
					UNTIL NOT again
					END_REPEAT;
				END_IF;
				// The writing end goes once no write is under way.
				IF CLOSE AND NOT closing THEN
					shut := TRUE;
				END_IF;
				closing := CLOSE;
				IF shut AND NOT BUSY THEN
					IF writable <> 0 THEN
						BYTES_STREAM_DROP_WRITABLE(stream := writable);
						writable := 0;
					END_IF;
					closed := TRUE;
					shut := FALSE;
				END_IF;
			END_FUNCTION_BLOCK

			/* Reads the value the future holds, which comes back after `DONE`. */
			{extern async 'wasi:cli/stdout@0.3.0' '[future-read-1]write-via-stream'}
			FUNCTION_BLOCK RESULT_FUTURE_READ
			VAR_INPUT
				future : UDINT;
			END_VAR
			VAR_OUTPUT
				DONE : BOOL;
				failed : BOOL;
				error : Wasi.Cli.Types.ERROR_CODE;
			END_VAR
			END_FUNCTION_BLOCK

			/* Lets go of the future's reading end, `future`. */
			{extern 'wasi:cli/stdout@0.3.0' '[future-drop-readable-1]write-via-stream'}
			FUNCTION RESULT_FUTURE_DROP_READABLE
			VAR_INPUT
				future : UDINT;
			END_VAR
			END_FUNCTION

			/* Reads the value the future holds, which comes back after `DONE`, then
			   lets go of the future's reading end: `future` is 0 from then on, and a
			   call with `future` 0 does nothing. */
			FUNCTION_BLOCK RESULT_FUTURE_GET
			VAR_IN_OUT
				future : UDINT;
			END_VAR
			VAR_OUTPUT
				DONE : BOOL;
				failed : BOOL;
				error : Wasi.Cli.Types.ERROR_CODE;
			END_VAR
			VAR
				call : RESULT_FUTURE_READ;
			END_VAR
				DONE := FALSE;
				IF future <> 0 THEN
					call(future := future);
					IF call.DONE THEN
						failed := call.failed;
						error := call.error;
						RESULT_FUTURE_DROP_READABLE(future := future);
						future := 0;
						DONE := TRUE;
					END_IF;
				END_IF;
			END_FUNCTION_BLOCK

			/* Writes text to `write-via-stream` through a stream of bytes it opens at
			   the first request. */
			FUNCTION_BLOCK WRITE_VIA_STREAM_WRITER
			VAR_INPUT
				/* A rising edge writes `IN`; the first opens the stream and calls
				   `write-via-stream` with it. An edge while `BUSY` is ignored. */
				REQ : BOOL;
				/* The text to write. */
				IN : STRING[4096];
				/* A rising edge ends the stream, once no write is under way. */
				CLOSE : BOOL;
			END_VAR
			VAR_OUTPUT
				/* TRUE while the reader has not taken all of `IN`. */
				BUSY : BOOL;
				/* TRUE in the call where the reader has taken all of `IN`, at once for an
				   empty text. */
				DONE : BOOL;
				/* TRUE once a write finds the reader gone, a request comes after `CLOSE`,
				   or the `result<_, error-code>` from `write-via-stream` is an error,
				   whose `error-code` is in `ERRORID`. */
				ERROR : BOOL;
				/* The `error-code` of the `result<_, error-code>` from `write-via-stream`,
				   when it is an error, which turns `ERROR` TRUE. */
				ERRORID : Wasi.Cli.Types.ERROR_CODE;
				/* TRUE once the `future<result<_, error-code>>` from `write-via-stream`
				   has its value. */
				ENDED : BOOL;
			END_VAR
			VAR
				open : BOOL;
				stream : BYTES_STREAM_WRITER;
				future : UDINT;
				answer : RESULT_FUTURE_GET;
			END_VAR
				// The stream, made at the first request and handed to the function.
				IF REQ AND NOT open THEN
					stream(REQ := FALSE, IN := IN, CLOSE := FALSE);
					future := Wasi.Cli.Stdout.WRITE_VIA_STREAM(data := stream.readable);
					open := TRUE;
				END_IF;
				IF open THEN
					stream(REQ := REQ, IN := IN, CLOSE := CLOSE);
					BUSY := stream.BUSY;
					DONE := stream.DONE;
					// The answer, read once it comes, and kept.
					answer(future := future);
					IF answer.DONE THEN
						ERRORID := answer.error;
						ENDED := TRUE;
					END_IF;
					ERROR := stream.ERROR OR answer.failed;
				END_IF;
			END_FUNCTION_BLOCK

			/* Writes bytes from an array to `write-via-stream` through a stream of
			   bytes it opens at the first request. */
			FUNCTION_BLOCK WRITE_VIA_STREAM_ARRAY_WRITER
			VAR_INPUT
				/* A rising edge writes the first `COUNT` bytes of `IN`; the first opens
				   the stream and calls `write-via-stream` with it. An edge while `BUSY` is
				   ignored. */
				REQ : BOOL;
				/* How many bytes of `IN` a request writes, from its first on. */
				COUNT : UDINT;
				/* A rising edge ends the stream, once no write is under way. */
				CLOSE : BOOL;
			END_VAR
			VAR_IN_OUT
				/* The bytes to write. The host reads them where they are while `BUSY`:
				   they stay as they are until `DONE`. */
				IN : ARRAY[*] OF BYTE;
			END_VAR
			VAR_OUTPUT
				/* TRUE while the reader has not taken all `COUNT` bytes. */
				BUSY : BOOL;
				/* TRUE in the call where the reader has taken all `COUNT` bytes, at once
				   for none. */
				DONE : BOOL;
				/* TRUE once a write finds the reader gone, a request comes after `CLOSE`,
				   or the `result<_, error-code>` from `write-via-stream` is an error,
				   whose `error-code` is in `ERRORID`. */
				ERROR : BOOL;
				/* The `error-code` of the `result<_, error-code>` from `write-via-stream`,
				   when it is an error, which turns `ERROR` TRUE. */
				ERRORID : Wasi.Cli.Types.ERROR_CODE;
				/* TRUE once the `future<result<_, error-code>>` from `write-via-stream`
				   has its value. */
				ENDED : BOOL;
			END_VAR
			VAR
				open : BOOL;
				stream : BYTES_STREAM_ARRAY_WRITER;
				future : UDINT;
				answer : RESULT_FUTURE_GET;
			END_VAR
				// The stream, made at the first request and handed to the function.
				IF REQ AND NOT open THEN
					stream(REQ := FALSE, COUNT := COUNT, CLOSE := FALSE, IN := IN);
					future := Wasi.Cli.Stdout.WRITE_VIA_STREAM(data := stream.readable);
					open := TRUE;
				END_IF;
				IF open THEN
					stream(REQ := REQ, COUNT := COUNT, CLOSE := CLOSE, IN := IN);
					BUSY := stream.BUSY;
					DONE := stream.DONE;
					// The answer, read once it comes, and kept.
					answer(future := future);
					IF answer.DONE THEN
						ERRORID := answer.error;
						ENDED := TRUE;
					END_IF;
					ERROR := stream.ERROR OR answer.failed;
				END_IF;
			END_FUNCTION_BLOCK
		END_NAMESPACE
	END_NAMESPACE
END_NAMESPACE
/* Not generated:
   - `BYTES_STREAM_CANCEL_WRITE`: a cancel blocks the scan.
   - `RESULT_FUTURE_CANCEL_READ`: a cancel blocks the scan. */

(* ---- wasi-clocks-monotonic-clock.st ---- *)
/* Generated from the WIT of wasi:clocks@0.3.0. DO NOT EDIT! */
NAMESPACE INTERNAL Wasi
	NAMESPACE Clocks
		/* WASI Monotonic Clock is a clock API intended to let users measure elapsed
		   time.

		   It is intended to be portable at least between Unix-family platforms and
		   Windows.

		   A monotonic clock is a clock which has an unspecified initial value, and
		   successive reads of the clock will produce non-decreasing values. */
		NAMESPACE MonotonicClock
			/* A mark on a monotonic clock is a number of nanoseconds since an
			   unspecified initial value, and can only be compared to instances from
			   the same monotonic-clock. */
			TYPE MARK : ULINT; END_TYPE

			/* Read the current value of the clock.

			   The clock is monotonic, therefore calling this function repeatedly will
			   produce a sequence of non-decreasing values.

			   For completeness, this function traps if it's not possible to represent
			   the value of the clock in a `mark`. Consequently, implementations
			   should ensure that the starting time is low enough to avoid the
			   possibility of overflow in practice. */
			{extern 'wasi:clocks/monotonic-clock@0.3.0' 'now'}
			FUNCTION NOW : MARK
			END_FUNCTION

			/* Query the resolution of the clock. Returns the duration of time
			   corresponding to a clock tick. */
			{extern 'wasi:clocks/monotonic-clock@0.3.0' 'get-resolution'}
			FUNCTION GET_RESOLUTION : Wasi.Clocks.Types.DURATION
			END_FUNCTION

			/* Wait until the specified mark has occurred. */
			{extern async 'wasi:clocks/monotonic-clock@0.3.0' 'wait-until'}
			FUNCTION_BLOCK WAIT_UNTIL
			VAR_INPUT
				when : MARK;
			END_VAR
			VAR_OUTPUT
				DONE : BOOL;
			END_VAR
			END_FUNCTION_BLOCK

			/* Wait for the specified duration to elapse. */
			{extern async 'wasi:clocks/monotonic-clock@0.3.0' 'wait-for'}
			FUNCTION_BLOCK WAIT_FOR
			VAR_INPUT
				how_long : Wasi.Clocks.Types.DURATION;
			END_VAR
			VAR_OUTPUT
				DONE : BOOL;
			END_VAR
			END_FUNCTION_BLOCK
		END_NAMESPACE
	END_NAMESPACE
END_NAMESPACE
